(*!
<summary>Selects the current stage of the independent runner contract suite.</summary>
*)
{attribute 'qualified_only'}
{attribute 'strict'}
TYPE TEST_RUNNER_CONTRACT_SCENARIO :
(
	STARTING,
	ELEMENT_TREE,
	CASE_ISOLATION,
	EMPTY_RUN,
	REPORTER_ABORT,
	DEADLINE,
	GROUP_TOPOLOGY,
	EXTERNAL_RECOVERY,
	DIAGNOSTICS,
	ADS_REPORTER_SUMMARY,
	ASSERTION_CONTRACTS,
	XML_ENCODING,
	RUNNER_TOPOLOGY,
	EXCEPTION_CLASSES,
	CONTEXT_OBJECTS,
	PATHS,
	INDEXED_CHILDREN,
	FINISHED
);
END_TYPE

(* stored: Version 1.1.0.1
   DUT TEST_RUNNER_CONTRACT_SCENARIO: Id {82985311-4b47-446a-aadf-00f6c9c896d9} *)
